(*
SPDX-FileCopyrightText: © 2026 Oleksandr Tiutyk <trofimich@gmail.com>
SPDX-License-Identifier: MIT
License: https://opensource.org/license/mit
*)

(*!
<summary>Exercises bounded multi-cycle completion and case-owned failure routing.</summary>
<description>
A nonzero Peer is failed during this body. Zero CompleteAfterCycle leaves completion to the deadline.
FailSelfWhileBusy asserts FALSE while returning TEST_CYCLE_RESULT.BUSY to verify immediate failure termination.
</description>
*)

{attribute 'no_explicit_call' := 'do not call this function block directly'}
FUNCTION_BLOCK AssertionIsolationProbe EXTENDS TOF_Testing.MultiCycleTest
VAR_INPUT
	Peer : POINTER TO AssertionIsolationProbe;
	UseDirectFailure : BOOL;
	FailSelfWhileBusy : BOOL;
	CompleteAfterCycle : UDINT := 3;
END_VAR
VAR_OUTPUT
	BodyCalls : UDINT;
	TeardownCalls : UDINT;
END_VAR
VAR_STAT
	//! <summary>Class name shared by all instances of this function block.</summary>
	{attribute 'hide'}
	_ClassName : STRING := __POUNAME();
END_VAR
VAR
	{attribute 'hide'}
	{attribute 'init_namespace'}
	_NamespaceName : STRING;
END_VAR

(*!
<summary>Resets per-run fixture observations.</summary>
*)
METHOD PROTECTED BeforeTest
BodyCalls := 0;
TeardownCalls := 0;
END_METHOD

(*!
<summary>Waits across scans or fails a peer and returns whether the scenario is done.</summary>
*)
METHOD PROTECTED ExecuteTest : TOF_Testing.TEST_CYCLE_RESULT
BodyCalls := BodyCalls + 1;

IF FailSelfWhileBusy THEN
	Assert.ThatBool(actual := FALSE).IsTrue();
	ExecuteTest := TOF_Testing.TEST_CYCLE_RESULT.BUSY;
ELSIF Peer <> 0 THEN
	Peer^.FailActiveCase(useDirectFailure := UseDirectFailure);
	ExecuteTest := TOF_Testing.TEST_CYCLE_RESULT.DONE;
ELSIF CompleteAfterCycle > TOF_Core.UnsignedInt32.ZERO AND_THEN CycleCount >= CompleteAfterCycle THEN
	Assert.ThatUDInt(actual := BodyCalls).ToBe(expected := CompleteAfterCycle);
	ExecuteTest := TOF_Testing.TEST_CYCLE_RESULT.DONE;
ELSE
	ExecuteTest := TOF_Testing.TEST_CYCLE_RESULT.BUSY;
END_IF
END_METHOD

(*!
<summary>Counts one cleanup for success, peer failure or timeout.</summary>
*)
METHOD PROTECTED AfterTest
TeardownCalls := TeardownCalls + 1;
END_METHOD

(*!
<summary>Reports through the receiving case while a different case is executing.</summary>
*)
METHOD INTERNAL FailActiveCase
VAR_INPUT
	useDirectFailure : BOOL;
END_VAR
IF useDirectFailure THEN
	RecordFailure(message := "Failure belongs to this case");
ELSE
	Assert.ThatBool(actual := FALSE).IsTrue();
END_IF
END_METHOD

//! <summary>Borrows the concrete class name for the lifetime of this instance; callers must not modify it.</summary>
{attribute 'monitoring' := 'call'}
PROPERTY ClassName : REFERENCE TO STRING
GET
ClassName REF= _ClassName;
END_GET
END_PROPERTY

//! <summary>Borrows the compiler-initialized namespace; callers must not modify the returned reference.</summary>
{attribute 'monitoring' := 'call'}
PROPERTY NamespaceName : REFERENCE TO STRING
GET
NamespaceName REF= _NamespaceName;
END_GET
END_PROPERTY

//! <summary>Reports the complete concrete instance size, excluding separately allocated storage.</summary>
{attribute 'monitoring' := 'call'}
PROPERTY SelfSize : ULINT
GET
SelfSize := XSIZEOF(THIS^);
END_GET
END_PROPERTY

END_FUNCTION_BLOCK

(* stored: Version 1.1.0.1
   POU AssertionIsolationProbe: Id {3b44f5d0-525a-4329-8d83-826a3b8a41f6}, SpecialFunc None
   Method BeforeTest: Id {4157ac7f-f099-49f0-afa6-036dd9820fa7}
   Method ExecuteTest: Id {ffa6eaa1-4c6d-4ab5-9e41-ae1a55d86fe3}
   Method AfterTest: Id {28bb19bb-0778-4688-8437-9611054e5f49}
   Method FailActiveCase: Id {a934b69f-fc76-4c33-8c45-a590b9139ed5}
   Property ClassName: Id {3be78a19-ae86-438c-bf68-ef66060a20f0}
   Get Get: Id {7fbdad64-e3ea-4e38-a958-a91ebe2bae00}
   Property NamespaceName: Id {5c3c7efe-619d-4b7c-818d-d108be261ac5}
   Get Get: Id {a72f69d0-618b-4fe8-90d7-02fa439d38a8}
   Property SelfSize: Id {557c3262-6b80-4782-b417-0607c92015f5}
   Get Get: Id {6b5d8f4e-9835-4be2-9b93-9cbce05eb119} *)
